(* IEC 61131-3 sources: codesys-framework/txt/application/WeVe Core (library)/60 Event/I_Event, 3 files *)

(* ---- Condition.method.st ---- *)
// Elke cyclus aanroepen voor een warning of alarm.
//   stijgende flank : event wordt actief en logt dat (met scPayload)
//   dalende flank   : logt dat de conditie weg is
//                     niet resetbaar -> event wordt meteen inactief
//                     resetbaar      -> event blijft actief tot Reset()
// Het event bouwt zelf de tekst op, de logger stuurt die alleen door.
// Geeft Active terug.
METHOD Condition : BOOL
VAR_INPUT
	xCondition 		: BOOL;
	scPayload 		: SC_EventPayload := (asPayload := [10('')]);	// mag weggelaten worden
END_VAR

(* ---- Log.method.st ---- *)
// Eenmalige melding, bv. drukknop of aanvraag. Logt OneShot, houdt geen toestand bij.
// TRUE = gelogd.
METHOD Log : BOOL
VAR_INPUT
	scPayload 		: SC_EventPayload := (asPayload := [10('')]);	// mag weggelaten worden
END_VAR

(* ---- Reset.method.st ---- *)
// Reset het event, maar enkel als de conditie weg is. Logt Reset.
// TRUE = event is niet (meer) actief.
METHOD Reset : BOOL
VAR_INPUT
END_VAR
